(* IEC 61131-3 sources: tsplc/packages/vscode-extension/tests/fixtures/build-tool/generated/types/ST_MotorZone, 3 files *)

(* ---- ST_MotorZone.st ---- *)
(*
Control signals and feedback for one 24 V motor-driven roller zone controller.
*)
TYPE ST_MotorZone :
STRUCT
	(* Normalized control signals toward one zone; mapping handles electrical polarity. *)
	Output : ST_MotorZoneOutput;
	(* Digital feedback from the zone controller, interpreted using the configured signal polarity. *)
	Input : ST_MotorZoneInput;
END_STRUCT
END_TYPE

(* ---- ST_MotorZoneInput.st ---- *)
(*
Control signals and feedback for one 24 V motor-driven roller zone controller.
*)
TYPE ST_MotorZoneInput :
STRUCT
	(* Zone sensor indication; TRUE when the photoeye is blocked. *)
	Sensor : BOOL;
	(* Aggregate error indication; no numeric diagnostic code is transmitted by this bit. *)
	Error : BOOL;
	(* Warning indication. *)
	Warning : BOOL;
	(* Synchronization indication; TRUE indicates motor running after polarity conversion. *)
	Sync : BOOL;
END_STRUCT
END_TYPE

(* ---- ST_MotorZoneOutput.st ---- *)
(*
Control signals and feedback for one 24 V motor-driven roller zone controller.
*)
TYPE ST_MotorZoneOutput :
STRUCT
	(* Run signal according to the configured zone mode. TRUE can force run or hold accumulation; FALSE can release accumulation. *)
	MotionAsserted : BOOL;
	(* Role depends on zone mode. Do not interpret as left/right sorter routing. *)
	DirectionOrSlaveErrorAsserted : BOOL;
	(* Optional speed reference in 0..10 V. Not metres/second and not a 4..20 mA signal. *)
	SpeedVolts : LREAL;
END_STRUCT
END_TYPE
